// TIA Portal V21 export
// export: Created 2026-11-11T00:48:10.6034942Z, ExportSetting WithDefaults, DisplayName Totally Integrated Automation Portal, DisplayVersion V21 Update 3, DisplayName STEP 7 Professional, DisplayVersion V21 Update 3, DisplayName STEP 7 Safety, DisplayVersion V21, DisplayName Tech WebApplication, DisplayVersion V21, DisplayName WinCC Basic/Comfort/Advanced, DisplayVersion V21 Update 3, DisplayName WinCC Unified, DisplayVersion V21 Update 3
FUNCTION_BLOCK "FB_Scl_sl016"   // FB30, SCL
{ S7_Optimized_Access := 'TRUE' }
VERSION : 0.1
// stored: AutoNumber true, IsIECCheckEnabled false, IsRetainMemResEnabled false, MemoryReserve 100, SetENOAutomatically false, UDAEnableTagReadback false
   VAR_INPUT
      v_cu : Bool;
      v_cd : Bool;
      v_r : Bool;
      v_ld : Bool;
      v_pv : Int;
   END_VAR
   VAR_OUTPUT
      v_qu : Bool;
      v_qd : Bool;
      v_cv : Char;
   END_VAR
   VAR
      inst { S7_SetPoint := 'True'} : CTUD_INT;
   END_VAR
BEGIN
   #inst(CU := #v_cu, CD := #v_cd, R := #v_r, LD := #v_ld, PV := #v_pv, QU => #v_qu, QD => #v_qd, CV => #v_cv);
END_FUNCTION_BLOCK
